FUNCTION "ROLL_PB21" : Void
{ S7_Optimized_Access := 'TRUE' }
VERSION : 0.1
VAR_TEMP
    r : Bool;
    a1 : Word;
    a2 : Word;
    activeDataBlock : Int;
    comparisonResults : Array[0..0] of Bool;
END_VAR
BEGIN
    #r := FALSE;
    #a1 := W#16#0000;
    #a2 := W#16#0000;
    #activeDataBlock := 0;
    // PB21, STEP 5 network 1
    #activeDataBlock := 15;
    // PB21, STEP 5 network 2
    #r := ((NOT "ROLL_IO".Input[3, 6]) AND (NOT "ROLL_State".M[13, 1]) AND (NOT "ROLL_State".M[5, 6]));
    "ROLL_State".M[99, 7] := #r;
    // PB21, STEP 5 network 3
    #r := ((NOT "ROLL_State".M[13, 3]) AND (NOT "ROLL_State".M[16, 6]) AND (NOT "ROLL_State".M[6, 0]) AND (NOT "ROLL_State".M[6, 2]) AND "ROLL_IO".Input[3, 0] AND "ROLL_IO".Input[5, 0] AND "ROLL_IO".Input[5, 2] AND "ROLL_IO".Input[5, 4]);
    "ROLL_State".M[100, 0] := #r;
    // PB21, STEP 5 network 4
    #r := "ROLL_State".M[190, 6];
    IF #r THEN "ROLL_State".M[100, 1] := TRUE; END_IF;
    #r := (((NOT "ROLL_State".M[190, 6]) AND "ROLL_IO".Input[5, 3]) OR (NOT "ROLL_IO".Input[0, 1]) OR (NOT "ROLL_State".M[0, 3]) OR (NOT "ROLL_State".M[100, 0]) OR "ROLL_State".M[190, 5]);
    IF #r THEN "ROLL_State".M[100, 1] := FALSE; END_IF;
    // PB21, STEP 5 network 5
    #r := "ROLL_State".M[190, 6];
    IF #r THEN "ROLL_State".M[100, 2] := TRUE; END_IF;
    #r := (("ROLL_IO".Input[5, 3] AND "ROLL_IO".Input[5, 6]) OR (NOT "ROLL_IO".Input[0, 1]) OR (NOT "ROLL_State".M[0, 3]) OR (NOT "ROLL_State".M[100, 0]) OR "ROLL_State".M[190, 5]);
    IF #r THEN "ROLL_State".M[100, 2] := FALSE; END_IF;
    // PB21, STEP 5 network 6
    #r := "ROLL_State".M[190, 6];
    IF #r THEN "ROLL_State".M[100, 3] := TRUE; END_IF;
    #r := (((NOT "ROLL_IO".Input[7, 5]) AND (NOT "ROLL_State".M[190, 6])) OR (NOT "ROLL_IO".Input[0, 1]) OR (NOT "ROLL_State".M[0, 3]) OR (NOT "ROLL_State".M[100, 0]) OR "ROLL_State".M[190, 5] OR "ROLL_State".M[5, 6] OR "ROLL_State".M[8, 5]);
    IF #r THEN "ROLL_State".M[100, 3] := FALSE; END_IF;
    // PB21, STEP 5 network 7
    #r := "ROLL_State".M[190, 6];
    IF #r THEN "ROLL_State".M[100, 4] := TRUE; END_IF;
    #r := (((NOT "ROLL_State".M[100, 0]) AND (NOT "ROLL_State".M[190, 6])) OR (NOT "ROLL_IO".Input[0, 1]) OR (NOT "ROLL_State".M[0, 3]) OR (NOT "ROLL_State".M[99, 7]) OR "ROLL_State".M[190, 5]);
    IF #r THEN "ROLL_State".M[100, 4] := FALSE; END_IF;
    // PB21, STEP 5 network 8
    #r := ((NOT "ROLL_State".M[31, 5]) AND (NOT "ROLL_State".M[5, 6]) AND ((NOT "ROLL_IO".Input[5, 6]) OR (NOT "ROLL_State".S5Timers[70].Q)) AND "ROLL_IO".Input[0, 2] AND "ROLL_IO".Input[3, 1] AND "ROLL_State".M[100, 0]);
    "ROLL_State".M[100, 5] := #r;
    // PB21, STEP 5 network 9
    #r := ((("ROLL_IO".Input[7, 5] AND "ROLL_State".S5Timers[97].Q) OR (NOT "ROLL_State".S5Timers[96].Q)) AND "ROLL_State".M[0, 3] AND "ROLL_State".M[100, 5]);
    "ROLL_State".M[100, 6] := #r;
    // PB21, STEP 5 network 10
    #r := ((((NOT "ROLL_IO".Input[7, 5]) AND "ROLL_State".S5Timers[96].Q) OR (NOT "ROLL_State".S5Timers[97].Q)) AND "ROLL_State".M[0, 3] AND "ROLL_State".M[100, 5]);
    "ROLL_State".M[100, 7] := #r;
    // PB21, STEP 5 network 11
    #r := "ROLL_State".M[190, 6];
    IF #r THEN "ROLL_State".M[101, 1] := TRUE; END_IF;
    #r := (((NOT "ROLL_State".M[190, 6]) AND "ROLL_IO".Input[5, 3] AND "ROLL_IO".Input[5, 6] AND "ROLL_IO".Input[6, 0]) OR (NOT "ROLL_IO".Input[0, 1]) OR (NOT "ROLL_State".M[0, 3]) OR (NOT "ROLL_State".M[100, 0]) OR "ROLL_State".M[190, 5]);
    IF #r THEN "ROLL_State".M[101, 1] := FALSE; END_IF;
    // PB21, STEP 5 network 12
    #r := "ROLL_State".M[190, 6];
    IF #r THEN "ROLL_State".M[101, 2] := TRUE; END_IF;
    #r := (((NOT "ROLL_State".M[190, 6]) AND "ROLL_IO".Input[5, 3] AND "ROLL_IO".Input[5, 6] AND "ROLL_IO".Input[6, 0]) OR (NOT "ROLL_IO".Input[0, 1]) OR (NOT "ROLL_State".M[0, 3]) OR (NOT "ROLL_State".M[100, 0]) OR "ROLL_State".M[190, 5]);
    IF #r THEN "ROLL_State".M[101, 2] := FALSE; END_IF;
    // PB21, STEP 5 network 13
    #r := "ROLL_State".M[190, 6];
    IF #r THEN "ROLL_State".M[101, 3] := TRUE; END_IF;
    #r := (((NOT "ROLL_State".M[190, 6]) AND ((NOT "ROLL_IO".Input[7, 5]) OR "ROLL_IO".Input[6, 0])) OR (NOT "ROLL_IO".Input[0, 1]) OR (NOT "ROLL_State".M[0, 3]) OR (NOT "ROLL_State".M[100, 0]) OR "ROLL_State".M[190, 5] OR "ROLL_State".M[5, 6] OR "ROLL_State".M[8, 5]);
    IF #r THEN "ROLL_State".M[101, 3] := FALSE; END_IF;
    // PB21, STEP 5 network 14
    #r := "ROLL_State".M[190, 6];
    IF #r THEN "ROLL_State".M[101, 4] := TRUE; END_IF;
    #r := (((NOT "ROLL_State".M[190, 6]) AND "ROLL_IO".Input[6, 0]) OR (NOT "ROLL_IO".Input[0, 1]) OR (NOT "ROLL_State".M[0, 3]) OR (NOT "ROLL_State".M[100, 0]) OR (NOT "ROLL_State".M[99, 7]) OR "ROLL_State".M[190, 5]);
    IF #r THEN "ROLL_State".M[101, 4] := FALSE; END_IF;
    // PB21, STEP 5 network 15
    #a2 := #a1;
    #a1 := W#16#2005;
    #r := "ROLL_IO".Input[6, 0];
    "ROLL_TimerOp"(Number := 121, Operation := 0, Signal := #r, Preset := #a1);
    // PB21, STEP 5 network 16
    #r := ((NOT "ROLL_State".M[31, 5]) AND (NOT "ROLL_State".M[5, 6]) AND (((NOT "ROLL_State".S5Timers[121].Q) AND "ROLL_State".M[101, 5]) OR (NOT "ROLL_IO".Input[6, 0])) AND "ROLL_IO".Input[0, 2] AND "ROLL_IO".Input[3, 1] AND "ROLL_State".M[100, 0]);
    "ROLL_State".M[101, 5] := #r;
    // PB21, STEP 5 network 17
    #r := ((("ROLL_IO".Input[7, 5] AND "ROLL_State".S5Timers[97].Q) OR (NOT "ROLL_State".S5Timers[96].Q)) AND "ROLL_State".M[101, 5]);
    "ROLL_State".M[101, 6] := #r;
    // PB21, STEP 5 network 18
    #r := ((((NOT "ROLL_IO".Input[7, 5]) AND "ROLL_State".S5Timers[96].Q) OR (NOT "ROLL_State".S5Timers[97].Q)) AND "ROLL_State".M[101, 5]);
    "ROLL_State".M[101, 7] := #r;
    // PB21, STEP 5 network 19
    #r := "ROLL_State".M[190, 6];
    IF #r THEN "ROLL_State".M[102, 1] := TRUE; END_IF;
    #r := (((NOT "ROLL_State".M[190, 6]) AND "ROLL_IO".Input[5, 3] AND "ROLL_IO".Input[5, 6] AND "ROLL_IO".Input[6, 0] AND "ROLL_IO".Input[6, 2]) OR (NOT "ROLL_IO".Input[0, 1]) OR (NOT "ROLL_State".M[0, 3]) OR (NOT "ROLL_State".M[100, 0]) OR "ROLL_State".M[190, 5]);
    IF #r THEN "ROLL_State".M[102, 1] := FALSE; END_IF;
    // PB21, STEP 5 network 20
    #r := "ROLL_State".M[190, 6];
    IF #r THEN "ROLL_State".M[102, 2] := TRUE; END_IF;
    #r := (((NOT "ROLL_State".M[190, 6]) AND "ROLL_IO".Input[6, 2]) OR (NOT "ROLL_IO".Input[0, 1]) OR (NOT "ROLL_State".M[0, 3]) OR (NOT "ROLL_State".M[100, 0]) OR "ROLL_State".M[190, 5]);
    IF #r THEN "ROLL_State".M[102, 2] := FALSE; END_IF;
    // PB21, STEP 5 network 21
    #r := "ROLL_State".M[190, 6];
    IF #r THEN "ROLL_State".M[102, 3] := TRUE; END_IF;
    #r := (((NOT "ROLL_State".M[190, 6]) AND ((NOT "ROLL_IO".Input[7, 5]) OR "ROLL_IO".Input[6, 2])) OR (NOT "ROLL_IO".Input[0, 1]) OR (NOT "ROLL_State".M[0, 3]) OR (NOT "ROLL_State".M[100, 0]) OR "ROLL_State".M[190, 5] OR "ROLL_State".M[5, 6] OR "ROLL_State".M[8, 5]);
    IF #r THEN "ROLL_State".M[102, 3] := FALSE; END_IF;
    // PB21, STEP 5 network 22
    #r := "ROLL_State".M[190, 6];
    IF #r THEN "ROLL_State".M[102, 4] := TRUE; END_IF;
    #r := (((NOT "ROLL_State".M[190, 6]) AND "ROLL_IO".Input[6, 2]) OR (NOT "ROLL_IO".Input[0, 1]) OR (NOT "ROLL_State".M[0, 3]) OR (NOT "ROLL_State".M[100, 0]) OR (NOT "ROLL_State".M[99, 7]) OR "ROLL_State".M[190, 5]);
    IF #r THEN "ROLL_State".M[102, 4] := FALSE; END_IF;
    // PB21, STEP 5 network 23
    #r := ((NOT "ROLL_State".M[31, 5]) AND (NOT "ROLL_State".M[5, 6]) AND (NOT "ROLL_State".S5Timers[72].Q) AND "ROLL_IO".Input[0, 2] AND "ROLL_IO".Input[3, 1] AND "ROLL_State".M[100, 0]);
    "ROLL_State".M[102, 5] := #r;
    // PB21, STEP 5 network 24
    #r := ((("ROLL_IO".Input[7, 5] AND "ROLL_State".S5Timers[97].Q) OR (NOT "ROLL_State".S5Timers[96].Q)) AND "ROLL_State".M[0, 3] AND "ROLL_State".M[102, 5]);
    "ROLL_State".M[102, 6] := #r;
    // PB21, STEP 5 network 25
    #r := ((((NOT "ROLL_IO".Input[7, 5]) AND "ROLL_State".S5Timers[96].Q) OR (NOT "ROLL_State".S5Timers[97].Q) OR "ROLL_State".M[0, 4]) AND "ROLL_State".M[102, 5]);
    "ROLL_State".M[102, 7] := #r;
    // PB21, STEP 5 network 26
    #r := "ROLL_State".M[190, 6];
    IF #r THEN "ROLL_State".M[105, 1] := TRUE; END_IF;
    #r := (((NOT "ROLL_State".M[190, 6]) AND "ROLL_State".M[0, 4]) OR (NOT "ROLL_IO".Input[0, 1]) OR (NOT "ROLL_State".M[0, 3]) OR (NOT "ROLL_State".M[100, 0]) OR "ROLL_State".M[190, 5]);
    IF #r THEN "ROLL_State".M[105, 1] := FALSE; END_IF;
    // PB21, STEP 5 network 27
    #r := "ROLL_State".M[190, 6];
    IF #r THEN "ROLL_State".M[105, 2] := TRUE; END_IF;
    #r := ((NOT "ROLL_IO".Input[0, 1]) OR (NOT "ROLL_State".M[0, 3]) OR (NOT "ROLL_State".M[100, 0]) OR "ROLL_IO".Input[6, 2] OR "ROLL_State".M[190, 5]);
    IF #r THEN "ROLL_State".M[105, 2] := FALSE; END_IF;
    // PB21, STEP 5 network 28
    #r := "ROLL_State".M[190, 6];
    IF #r THEN "ROLL_State".M[105, 3] := TRUE; END_IF;
    #r := (((NOT "ROLL_State".M[190, 6]) AND ((NOT "ROLL_IO".Input[7, 5]) OR "ROLL_State".M[0, 4])) OR (NOT "ROLL_IO".Input[0, 1]) OR (NOT "ROLL_State".M[0, 3]) OR (NOT "ROLL_State".M[100, 0]) OR "ROLL_State".M[190, 5] OR "ROLL_State".M[5, 6] OR "ROLL_State".M[8, 5]);
    IF #r THEN "ROLL_State".M[105, 3] := FALSE; END_IF;
    // PB21, STEP 5 network 29
    #r := "ROLL_State".M[190, 6];
    IF #r THEN "ROLL_State".M[105, 4] := TRUE; END_IF;
    #r := (((NOT "ROLL_State".M[190, 6]) AND "ROLL_State".M[0, 4]) OR (NOT "ROLL_IO".Input[0, 1]) OR (NOT "ROLL_State".M[0, 3]) OR (NOT "ROLL_State".M[100, 0]) OR (NOT "ROLL_State".M[99, 7]) OR "ROLL_State".M[190, 5]);
    IF #r THEN "ROLL_State".M[105, 4] := FALSE; END_IF;
    // PB21, STEP 5 network 30
    #a2 := #a1;
    #a1 := W#16#2005;
    #r := "ROLL_State".M[0, 4];
    "ROLL_TimerOp"(Number := 120, Operation := 0, Signal := #r, Preset := #a1);
    // PB21, STEP 5 network 31
    #r := ((NOT "ROLL_State".M[31, 5]) AND (NOT "ROLL_State".M[5, 6]) AND (((NOT "ROLL_State".S5Timers[120].Q) AND "ROLL_State".M[105, 5]) OR (NOT "ROLL_State".M[0, 4])) AND "ROLL_IO".Input[0, 2] AND "ROLL_IO".Input[3, 1] AND "ROLL_State".M[100, 0]);
    "ROLL_State".M[105, 5] := #r;
    // PB21, STEP 5 network 32
    #r := ((("ROLL_IO".Input[7, 5] AND "ROLL_State".S5Timers[97].Q) OR (NOT "ROLL_State".S5Timers[96].Q)) AND "ROLL_State".M[105, 5]);
    "ROLL_State".M[105, 6] := #r;
    // PB21, STEP 5 network 33
    #r := ((((NOT "ROLL_IO".Input[7, 5]) AND "ROLL_State".S5Timers[96].Q) OR (NOT "ROLL_State".S5Timers[97].Q)) AND "ROLL_State".M[105, 5]);
    "ROLL_State".M[105, 7] := #r;
    // PB21, STEP 5 network 34
    #r := ((((NOT "ROLL_IO".Input[5, 5]) AND ("ROLL_State".M[40, 5] OR "ROLL_State".M[42, 1]) AND "ROLL_State".M[31, 5]) OR (NOT "ROLL_IO".Input[5, 6])) AND "ROLL_IO".Input[0, 2] AND "ROLL_IO".Input[3, 1] AND "ROLL_State".M[100, 0]);
    "ROLL_State".M[103, 0] := #r;
    // PB21, STEP 5 network 35
    #r := (((NOT "ROLL_IO".Input[5, 3]) OR (NOT "ROLL_IO".Input[6, 0]) OR (NOT "ROLL_State".S5Timers[121].Q)) AND "ROLL_IO".Input[3, 1] AND "ROLL_State".M[100, 0] AND "ROLL_State".M[31, 5]);
    "ROLL_State".M[103, 3] := #r;
    // PB21, STEP 5 network 36
    #r := (((NOT "ROLL_IO".Input[5, 6]) AND "ROLL_IO".Input[0, 2]) OR (("ROLL_State".M[103, 0] OR "ROLL_State".M[103, 3]) AND "ROLL_State".S5Timers[62].Q AND "ROLL_State".S5Timers[97].Q));
    "ROLL_State".M[103, 1] := #r;
    // PB21, STEP 5 network 37
    #r := ((NOT "ROLL_IO".Input[6, 2]) AND "ROLL_IO".Input[3, 1] AND "ROLL_State".M[100, 0] AND "ROLL_State".M[31, 5]);
    "ROLL_State".M[103, 4] := #r;
    // PB21, STEP 5 network 38
    #a2 := #a1;
    #a1 := W#16#1050;
    #r := ("ROLL_IO".Output[22, 3] AND "ROLL_State".M[103, 4]);
    "ROLL_TimerOp"(Number := 119, Operation := 1, Signal := #r, Preset := #a1);
    // PB21, STEP 5 network 39
    #r := (((("ROLL_State".M[103, 0] OR "ROLL_State".M[103, 3]) AND "ROLL_State".S5Timers[96].Q) OR "ROLL_State".M[103, 4] OR "ROLL_State".S5Timers[119].Q) AND "ROLL_State".S5Timers[62].Q);
    "ROLL_State".M[103, 2] := #r;
    // PB21, STEP 5 network 40
    #r := "ROLL_State".M[190, 6];
    IF #r THEN "ROLL_State".M[104, 0] := TRUE; END_IF;
    #r := (((NOT "ROLL_State".M[190, 6]) AND ((NOT "ROLL_IO".Input[5, 0]) OR (NOT "ROLL_IO".Input[5, 2]) OR (NOT "ROLL_IO".Input[5, 4]))) OR (NOT "ROLL_IO".Input[0, 1]) OR (NOT "ROLL_IO".Input[7, 0]) OR (NOT "ROLL_State".M[26, 5]) OR (NOT "ROLL_State".M[99, 7]) OR "ROLL_State".M[16, 6] OR "ROLL_State".M[190, 5]);
    IF #r THEN "ROLL_State".M[104, 0] := FALSE; END_IF;
    // PB21, STEP 5 network 41
    #r := "ROLL_State".M[190, 6];
    IF #r THEN "ROLL_State".M[104, 1] := TRUE; END_IF;
    #r := (((NOT "ROLL_State".M[190, 6]) AND ((NOT "ROLL_IO".Input[5, 0]) OR (NOT "ROLL_IO".Input[5, 2]) OR (NOT "ROLL_IO".Input[5, 4]))) OR (NOT "ROLL_IO".Input[0, 1]) OR (NOT "ROLL_State".M[26, 0]) OR (NOT "ROLL_State".M[99, 7]) OR "ROLL_State".M[16, 6] OR "ROLL_State".M[190, 5]);
    IF #r THEN "ROLL_State".M[104, 1] := FALSE; END_IF;
    // PB21, STEP 5 network 42
    #r := "ROLL_State".M[190, 6];
    IF #r THEN "ROLL_State".M[104, 4] := TRUE; END_IF;
    #r := (((NOT "ROLL_State".M[190, 6]) AND ((NOT "ROLL_IO".Input[5, 0]) OR (NOT "ROLL_IO".Input[5, 2]) OR (NOT "ROLL_IO".Input[5, 4]))) OR (NOT "ROLL_IO".Input[0, 1]) OR (NOT "ROLL_IO".Input[4, 7]) OR (NOT "ROLL_State".M[27, 4]) OR (NOT "ROLL_State".M[99, 7]) OR "ROLL_State".M[16, 6] OR "ROLL_State".M[190, 5]);
    IF #r THEN "ROLL_State".M[104, 4] := FALSE; END_IF;
    // PB21, STEP 5 network 43
    #r := "ROLL_State".M[190, 6];
    IF #r THEN "ROLL_State".M[104, 5] := TRUE; END_IF;
    #r := (((NOT "ROLL_State".M[190, 6]) AND "ROLL_IO".Input[5, 3] AND "ROLL_IO".Input[5, 6] AND "ROLL_IO".Input[6, 0] AND "ROLL_IO".Input[6, 2]) OR (NOT "ROLL_IO".Input[0, 1]) OR (NOT "ROLL_State".M[100, 0]) OR (NOT "ROLL_State".M[24, 1]) OR "ROLL_State".M[190, 5]);
    IF #r THEN "ROLL_State".M[104, 5] := FALSE; END_IF;
    // PB21, STEP 5 network 44
    #r := "ROLL_State".M[190, 6];
    IF #r THEN "ROLL_State".M[104, 6] := TRUE; END_IF;
    #r := (((NOT "ROLL_State".M[190, 6]) AND (("ROLL_IO".Input[5, 3] AND "ROLL_IO".Input[5, 6] AND "ROLL_IO".Input[6, 0]) OR (NOT "ROLL_IO".Input[7, 5]))) OR (NOT "ROLL_IO".Input[0, 1]) OR (NOT "ROLL_State".M[100, 0]) OR (NOT "ROLL_State".M[25, 0]) OR "ROLL_State".M[190, 5] OR "ROLL_State".M[5, 6] OR "ROLL_State".M[8, 5]);
    IF #r THEN "ROLL_State".M[104, 6] := FALSE; END_IF;
    // PB21, STEP 5 network 45
    #r := "ROLL_State".S5Timers[59].Q;
    "ROLL_IO".Output[17, 0] := #r;
    // PB21, STEP 5 network 46
    #r := ("ROLL_IO".Input[6, 5] AND "ROLL_State".M[100, 0]);
    "ROLL_IO".Output[17, 5] := #r;
    RETURN;
END_FUNCTION

FUNCTION "ROLL_PB23" : Void
{ S7_Optimized_Access := 'TRUE' }
VERSION : 0.1
VAR_TEMP
    r : Bool;
    a1 : Word;
    a2 : Word;
    activeDataBlock : Int;
    comparisonResults : Array[0..0] of Bool;
END_VAR
BEGIN
    #r := FALSE;
    #a1 := W#16#0000;
    #a2 := W#16#0000;
    #activeDataBlock := 0;
    // PB23, STEP 5 network 1
    #activeDataBlock := 15;
    // PB23, STEP 5 network 2
    #r := (("ROLL_State".M[40, 3] OR "ROLL_State".M[40, 4] OR "ROLL_State".M[40, 5]) AND "ROLL_State".M[111, 4]);
    "ROLL_State".M[240, 0] := #r;
    // PB23, STEP 5 network 3
    #a2 := #a1;
    #a1 := W#16#2120;
    #r := "ROLL_State".M[240, 0];
    "ROLL_TimerOp"(Number := 51, Operation := 1, Signal := #r, Preset := #a1);
    #r := "ROLL_State".S5Timers[51].Q;
    "ROLL_IO".Output[19, 0] := #r;
    // PB23, STEP 5 network 4
    #a2 := #a1;
    #a1 := W#16#1050;
    #r := ((NOT "ROLL_State".M[6, 1]) AND ("ROLL_State".M[40, 4] OR "ROLL_State".M[40, 5]) AND "ROLL_IO".Output[19, 0] AND "ROLL_State".M[240, 0] AND "ROLL_State".M[35, 2] AND "ROLL_State".S5Timers[70].Q);
    "ROLL_TimerOp"(Number := 52, Operation := 0, Signal := #r, Preset := #a1);
    #r := "ROLL_State".S5Timers[52].Q;
    "ROLL_IO".Output[19, 1] := #r;
    // PB23, STEP 5 network 5
    #r := ("ROLL_IO".Input[0, 2] AND "ROLL_IO".Input[0, 4]);
    IF #r THEN "ROLL_State".M[103, 7] := TRUE; END_IF;
    #r := (NOT "ROLL_State".S5Timers[59].Q);
    IF #r THEN "ROLL_State".M[103, 7] := FALSE; END_IF;
    // PB23, STEP 5 network 6
    #a2 := #a1;
    #a1 := W#16#3360;
    #r := "ROLL_State".S5Timers[59].Q;
    "ROLL_TimerOp"(Number := 76, Operation := 0, Signal := #r, Preset := #a1);
    // PB23, STEP 5 network 7
    #r := ((NOT "ROLL_State".M[13, 3]) AND (NOT "ROLL_State".M[5, 6]) AND (NOT "ROLL_State".M[6, 2]) AND (NOT "ROLL_State".M[6, 3]) AND (((NOT "ROLL_State".S5Timers[76].Q) AND "ROLL_IO".Input[2, 2]) OR "ROLL_State".M[103, 7] OR "ROLL_State".M[152, 0]) AND ("ROLL_IO".Input[2, 2] OR "ROLL_State".M[152, 0]) AND "ROLL_IO".Input[3, 4] AND "ROLL_IO".Input[5, 6] AND "ROLL_State".S5Timers[59].Q);
    "ROLL_IO".Output[19, 5] := #r;
    // PB23, STEP 5 network 8
    #r := ((NOT "ROLL_State".M[5, 6]) AND (NOT "ROLL_State".M[6, 1]) AND ("ROLL_IO".Input[0, 1] OR "ROLL_IO".Input[0, 2]) AND "ROLL_IO".Input[3, 1] AND "ROLL_IO".Input[3, 4] AND "ROLL_State".M[0, 3] AND "ROLL_State".M[100, 0] AND "ROLL_State".S5Timers[70].Q);
    "ROLL_State".M[240, 0] := #r;
    // PB23, STEP 5 network 9
    #r := ((NOT "ROLL_IO".Output[20, 6]) AND (NOT "ROLL_State".M[5, 6]) AND (NOT "ROLL_State".M[8, 5]) AND (NOT "ROLL_State".S5Timers[96].Q) AND (("ROLL_State".M[100, 0] AND "ROLL_State".M[103, 1]) OR "ROLL_State".M[102, 6] OR "ROLL_State".M[104, 6]));
    "ROLL_IO".Output[20, 4] := #r;
    "ROLL_IO".Output[22, 6] := #r;
    // PB23, STEP 5 network 10
    #r := ((NOT "ROLL_IO".Output[20, 1]) AND ("ROLL_State".M[104, 0] OR "ROLL_State".M[104, 1] OR "ROLL_State".M[104, 4] OR "ROLL_State".M[152, 1]) AND "ROLL_State".M[99, 7]);
    "ROLL_IO".Output[20, 6] := #r;
    // PB23, STEP 5 network 11
    #r := ("ROLL_State".M[102, 7] OR "ROLL_State".M[103, 2] OR "ROLL_State".M[104, 5]);
    "ROLL_State".M[240, 0] := #r;
    // PB23, STEP 5 network 12
    #r := ((NOT "ROLL_State".M[13, 4]) AND (NOT "ROLL_State".M[6, 0]) AND (NOT "ROLL_State".M[6, 2]) AND (NOT "ROLL_State".M[7, 7]) AND "ROLL_IO".Input[3, 1] AND "ROLL_IO".Input[5, 0] AND "ROLL_IO".Input[5, 2] AND "ROLL_IO".Input[5, 4] AND "ROLL_State".M[240, 0]);
    "ROLL_IO".Output[20, 1] := #r;
    // PB23, STEP 5 network 13
    #r := "ROLL_State".M[103, 1];
    "ROLL_IO".Output[22, 2] := #r;
    // PB23, STEP 5 network 14
    #r := ("ROLL_State".M[102, 1] OR "ROLL_State".M[102, 2] OR "ROLL_State".M[102, 3] OR "ROLL_State".M[102, 6] OR "ROLL_State".M[102, 7] OR "ROLL_State".M[103, 2]);
    "ROLL_IO".Output[22, 3] := #r;
    // PB23, STEP 5 network 15
    #r := "ROLL_State".S5Timers[85].Q;
    "ROLL_IO".Output[21, 3] := #r;
    // PB23, STEP 5 network 16
    #a2 := #a1;
    #a1 := W#16#1020;
    #r := "ROLL_IO".Output[20, 6];
    "ROLL_TimerOp"(Number := 47, Operation := 1, Signal := #r, Preset := #a1);
    // PB23, STEP 5 network 17
    #r := ((NOT "ROLL_IO".Output[21, 5]) AND (NOT "ROLL_IO".Output[22, 3]) AND (NOT "ROLL_IO".Output[22, 6]) AND (("ROLL_IO".Output[21, 4] AND "ROLL_State".S5Timers[47].Q) OR "ROLL_State".M[104, 0] OR "ROLL_State".M[152, 1]));
    "ROLL_IO".Output[21, 4] := #r;
    // PB23, STEP 5 network 18
    #r := ((NOT "ROLL_IO".Output[21, 4]) AND "ROLL_State".M[152, 0]);
    "ROLL_IO".Output[21, 5] := #r;
    // PB23, STEP 5 network 19
    RETURN;
END_FUNCTION

FUNCTION "ROLL_PB24" : Void
{ S7_Optimized_Access := 'TRUE' }
VERSION : 0.1
VAR_TEMP
    r : Bool;
    a1 : Word;
    a2 : Word;
    activeDataBlock : Int;
    comparisonResults : Array[0..0] of Bool;
END_VAR
BEGIN
    #r := FALSE;
    #a1 := W#16#0000;
    #a2 := W#16#0000;
    #activeDataBlock := 0;
    // PB24, STEP 5 network 1
    #activeDataBlock := 15;
    // PB24, STEP 5 network 2
    #r := ("ROLL_IO".Input[5, 0] AND "ROLL_State".M[13, 3] AND "ROLL_State".S5Timers[59].Q);
    "ROLL_State".M[240, 0] := #r;
    // PB24, STEP 5 network 3
    #a2 := #a1;
    #a1 := "ROLL_GetDW"(DbNumber := #activeDataBlock, Index := 54);
    #r := (NOT "ROLL_State".S5Timers[53].Q);
    "ROLL_TimerOp"(Number := 54, Operation := 0, Signal := #r, Preset := #a1);
    #a2 := #a1;
    #a1 := "ROLL_GetDW"(DbNumber := #activeDataBlock, Index := 53);
    #r := "ROLL_State".S5Timers[54].Q;
    "ROLL_TimerOp"(Number := 53, Operation := 1, Signal := #r, Preset := #a1);
    #r := "ROLL_State".M[240, 0];
    "ROLL_TimerOp"(Number := 53, Operation := 2, Signal := #r, Preset := #a1);
    #r := ((NOT "ROLL_State".M[40, 5]) AND "ROLL_State".S5Timers[53].Q);
    "ROLL_IO".Output[19, 4] := #r;
    // PB24, STEP 5 network 4
    RETURN;
END_FUNCTION

FUNCTION "ROLL_PB25" : Void
{ S7_Optimized_Access := 'TRUE' }
VERSION : 0.1
VAR_TEMP
    r : Bool;
    a1 : Word;
    a2 : Word;
    activeDataBlock : Int;
    comparisonResults : Array[0..14] of Bool;
END_VAR
BEGIN
    #r := FALSE;
    #a1 := W#16#0000;
    #a2 := W#16#0000;
    #activeDataBlock := 0;
    // PB25, STEP 5 network 1
    #activeDataBlock := 15;
    // PB25, STEP 5 network 2
    #a2 := #a1;
    #a1 := "ROLL_GetM"(FirstByte := 5, Width := 8);
    #a2 := #a1;
    #a1 := W#16#0000;
    #comparisonResults[0] := (WORD_TO_INT(#a2) <> WORD_TO_INT(#a1));
    #r := #comparisonResults[0];
    "ROLL_State".M[87, 0] := #r;
    // PB25, STEP 5 network 3
    #a2 := #a1;
    #a1 := "ROLL_GetM"(FirstByte := 6, Width := 8);
    #a2 := #a1;
    #a1 := W#16#0000;
    #comparisonResults[1] := (WORD_TO_INT(#a2) <> WORD_TO_INT(#a1));
    #r := #comparisonResults[1];
    "ROLL_State".M[87, 1] := #r;
    // PB25, STEP 5 network 4
    #a2 := #a1;
    #a1 := "ROLL_GetM"(FirstByte := 7, Width := 8);
    #a2 := #a1;
    #a1 := W#16#0000;
    #comparisonResults[2] := (WORD_TO_INT(#a2) <> WORD_TO_INT(#a1));
    #r := #comparisonResults[2];
    "ROLL_State".M[87, 2] := #r;
    // PB25, STEP 5 network 5
    #a2 := #a1;
    #a1 := "ROLL_GetM"(FirstByte := 8, Width := 8);
    #a2 := #a1;
    #a1 := W#16#0000;
    #comparisonResults[3] := (WORD_TO_INT(#a2) <> WORD_TO_INT(#a1));
    #r := #comparisonResults[3];
    "ROLL_State".M[87, 3] := #r;
    // PB25, STEP 5 network 6
    #a2 := #a1;
    #a1 := "ROLL_GetM"(FirstByte := 9, Width := 8);
    #a2 := #a1;
    #a1 := W#16#0000;
    #comparisonResults[4] := (WORD_TO_INT(#a2) <> WORD_TO_INT(#a1));
    #r := #comparisonResults[4];
    "ROLL_State".M[87, 4] := #r;
    // PB25, STEP 5 network 7
    #a2 := #a1;
    #a1 := "ROLL_GetM"(FirstByte := 10, Width := 8);
    #a2 := #a1;
    #a1 := W#16#0000;
    #comparisonResults[5] := (WORD_TO_INT(#a2) <> WORD_TO_INT(#a1));
    #r := #comparisonResults[5];
    "ROLL_State".M[87, 5] := #r;
    // PB25, STEP 5 network 8
    #a2 := #a1;
    #a1 := "ROLL_GetM"(FirstByte := 11, Width := 8);
    #a2 := #a1;
    #a1 := W#16#0000;
    #comparisonResults[6] := (WORD_TO_INT(#a2) <> WORD_TO_INT(#a1));
    #r := #comparisonResults[6];
    "ROLL_State".M[87, 6] := #r;
    // PB25, STEP 5 network 9
    #a2 := #a1;
    #a1 := "ROLL_GetM"(FirstByte := 12, Width := 8);
    #a2 := #a1;
    #a1 := W#16#0000;
    #comparisonResults[7] := (WORD_TO_INT(#a2) <> WORD_TO_INT(#a1));
    #r := #comparisonResults[7];
    "ROLL_State".M[87, 7] := #r;
    // PB25, STEP 5 network 10
    #a2 := #a1;
    #a1 := "ROLL_GetM"(FirstByte := 13, Width := 8);
    #a2 := #a1;
    #a1 := W#16#0000;
    #comparisonResults[8] := (WORD_TO_INT(#a2) <> WORD_TO_INT(#a1));
    #r := #comparisonResults[8];
    "ROLL_State".M[88, 0] := #r;
    // PB25, STEP 5 network 11
    #a2 := #a1;
    #a1 := "ROLL_GetM"(FirstByte := 14, Width := 8);
    #a2 := #a1;
    #a1 := W#16#0000;
    #comparisonResults[9] := (WORD_TO_INT(#a2) <> WORD_TO_INT(#a1));
    #r := #comparisonResults[9];
    "ROLL_State".M[88, 1] := #r;
    // PB25, STEP 5 network 12
    #a2 := #a1;
    #a1 := "ROLL_GetM"(FirstByte := 15, Width := 8);
    #a2 := #a1;
    #a1 := W#16#0000;
    #comparisonResults[10] := (WORD_TO_INT(#a2) <> WORD_TO_INT(#a1));
    #r := #comparisonResults[10];
    "ROLL_State".M[88, 2] := #r;
    // PB25, STEP 5 network 13
    #a2 := #a1;
    #a1 := "ROLL_GetM"(FirstByte := 16, Width := 8);
    #a2 := #a1;
    #a1 := W#16#0000;
    #comparisonResults[11] := (WORD_TO_INT(#a2) <> WORD_TO_INT(#a1));
    #r := #comparisonResults[11];
    "ROLL_State".M[88, 3] := #r;
    // PB25, STEP 5 network 14
    #a2 := #a1;
    #a1 := "ROLL_GetM"(FirstByte := 17, Width := 8);
    #a2 := #a1;
    #a1 := W#16#0000;
    #comparisonResults[12] := (WORD_TO_INT(#a2) <> WORD_TO_INT(#a1));
    #r := #comparisonResults[12];
    "ROLL_State".M[88, 4] := #r;
    // PB25, STEP 5 network 15
    #a2 := #a1;
    #a1 := "ROLL_GetM"(FirstByte := 18, Width := 8);
    #a2 := #a1;
    #a1 := W#16#0000;
    #comparisonResults[13] := (WORD_TO_INT(#a2) <> WORD_TO_INT(#a1));
    #r := #comparisonResults[13];
    "ROLL_State".M[88, 5] := #r;
    // PB25, STEP 5 network 16
    #a2 := #a1;
    #a1 := "ROLL_GetM"(FirstByte := 19, Width := 8);
    #a2 := #a1;
    #a1 := W#16#0000;
    #comparisonResults[14] := (WORD_TO_INT(#a2) <> WORD_TO_INT(#a1));
    #r := #comparisonResults[14];
    "ROLL_State".M[88, 6] := #r;
    // PB25, STEP 5 network 17
    #r := ("ROLL_State".M[87, 0] OR "ROLL_State".M[87, 1] OR "ROLL_State".M[87, 2] OR "ROLL_State".M[87, 3] OR "ROLL_State".M[87, 4] OR "ROLL_State".M[87, 5] OR "ROLL_State".M[87, 6] OR "ROLL_State".M[87, 7] OR "ROLL_State".M[88, 0] OR "ROLL_State".M[88, 1] OR "ROLL_State".M[88, 2] OR "ROLL_State".M[88, 3] OR "ROLL_State".M[88, 4] OR "ROLL_State".M[88, 5] OR "ROLL_State".M[88, 6]);
    "ROLL_State".M[88, 7] := #r;
    // PB25, STEP 5 network 18
    #r := ("ROLL_IO".Input[1, 2] OR "ROLL_State".M[88, 7]);
    "ROLL_IO".Output[16, 4] := #r;
    // PB25, STEP 5 network 19
    #r := (("ROLL_State".M[3, 6] AND "ROLL_State".M[31, 6]) OR "ROLL_IO".Input[1, 2]);
    "ROLL_IO".Output[16, 5] := #r;
    // PB25, STEP 5 network 20
    #r := ("ROLL_IO".Input[1, 2] OR "ROLL_IO".Input[3, 4]);
    "ROLL_IO".Output[16, 0] := #r;
    // PB25, STEP 5 network 21
    #r := (((NOT "ROLL_State".M[31, 5]) AND "ROLL_State".M[28, 4]) OR ("ROLL_State".M[3, 6] AND "ROLL_State".M[74, 0]) OR "ROLL_IO".Input[1, 2]);
    "ROLL_IO".Output[16, 2] := #r;
    // PB25, STEP 5 network 22
    #r := (("ROLL_State".M[3, 6] AND "ROLL_State".M[31, 5]) OR "ROLL_IO".Input[1, 2] OR "ROLL_State".M[31, 4]);
    "ROLL_IO".Output[16, 3] := #r;
    // PB25, STEP 5 network 23
    #r := "ROLL_IO".Input[2, 0];
    "ROLL_IO".Output[19, 3] := #r;
    // PB25, STEP 5 network 24
    #r := (((("ROLL_IO".Input[14, 0] AND "ROLL_State".M[37, 1]) OR "ROLL_State".M[53, 6]) AND "ROLL_IO".Input[0, 2]) OR ("ROLL_IO".Input[0, 1] AND "ROLL_State".M[190, 6] AND "ROLL_State".M[20, 7]));
    IF #r THEN "ROLL_State".M[71, 5] := TRUE; END_IF;
    #r := (("ROLL_IO".Input[0, 1] AND "ROLL_State".M[190, 5] AND "ROLL_State".M[20, 7]) OR ("ROLL_IO".Input[0, 2] AND "ROLL_State".M[37, 2]));
    IF #r THEN "ROLL_State".M[71, 5] := FALSE; END_IF;
    #r := "ROLL_State".M[71, 5];
    "ROLL_IO".Output[17, 7] := #r;
    // PB25, STEP 5 network 25
    RETURN;
END_FUNCTION

FUNCTION "ROLL_PB50" : Void
{ S7_Optimized_Access := 'TRUE' }
VERSION : 0.1
VAR_TEMP
    r : Bool;
    a1 : Word;
    a2 : Word;
    activeDataBlock : Int;
    comparisonResults : Array[0..0] of Bool;
END_VAR
BEGIN
    #r := FALSE;
    #a1 := W#16#0000;
    #a2 := W#16#0000;
    #activeDataBlock := 0;
    // PB50, STEP 5 network 1
    #activeDataBlock := 15;
    // PB50, STEP 5 network 2
    #r := "ROLL_State".M[0, 1];
    IF #r THEN "ROLL_State".M[0, 2] := FALSE; END_IF;
    // PB50, STEP 5 network 3
    #a2 := #a1;
    #a1 := W#16#2008;
    #r := ((NOT "ROLL_State".M[0, 1]) AND "ROLL_IO".Input[3, 0]);
    "ROLL_TimerOp"(Number := 11, Operation := 0, Signal := #r, Preset := #a1);
    // PB50, STEP 5 network 4
    #a2 := #a1;
    #a1 := W#16#1020;
    #r := "ROLL_State".M[29, 0];
    "ROLL_TimerOp"(Number := 13, Operation := 0, Signal := #r, Preset := #a1);
    // PB50, STEP 5 network 5
    RETURN;
END_FUNCTION

FUNCTION "ROLL_PB51" : Void
{ S7_Optimized_Access := 'TRUE' }
VERSION : 0.1
VAR_TEMP
    r : Bool;
    a1 : Word;
    a2 : Word;
    activeDataBlock : Int;
    comparisonResults : Array[0..0] of Bool;
END_VAR
BEGIN
    #r := FALSE;
    #a1 := W#16#0000;
    #a2 := W#16#0000;
    #activeDataBlock := 0;
    // PB51, STEP 5 network 1
    #a2 := #a1;
    #a1 := W#16#2060;
    #r := "ROLL_IO".Output[24, 0];
    "ROLL_TimerOp"(Number := 15, Operation := 0, Signal := #r, Preset := #a1);
    // PB51, STEP 5 network 2
    #a2 := #a1;
    #a1 := W#16#3360;
    #r := ((NOT "ROLL_IO".Input[5, 6]) AND "ROLL_State".M[31, 5]);
    "ROLL_TimerOp"(Number := 16, Operation := 0, Signal := #r, Preset := #a1);
    // PB51, STEP 5 network 3
    #a2 := #a1;
    #a1 := W#16#1010;
    #r := "ROLL_State".M[37, 5];
    "ROLL_TimerOp"(Number := 18, Operation := 0, Signal := #r, Preset := #a1);
    // PB51, STEP 5 network 4
    #a2 := #a1;
    #a1 := W#16#2015;
    #r := (((NOT "ROLL_IO".Input[124, 1]) AND "ROLL_IO".Output[112, 1]) OR ((NOT "ROLL_IO".Input[124, 2]) AND "ROLL_IO".Output[112, 2]));
    "ROLL_TimerOp"(Number := 19, Operation := 0, Signal := #r, Preset := #a1);
    // PB51, STEP 5 network 5
    #a2 := #a1;
    #a1 := W#16#1010;
    #r := (("ROLL_IO".Input[123, 4] OR "ROLL_IO".Input[123, 5]) AND "ROLL_IO".Output[112, 0]);
    "ROLL_TimerOp"(Number := 20, Operation := 0, Signal := #r, Preset := #a1);
    // PB51, STEP 5 network 6
    #a2 := #a1;
    #a1 := W#16#1050;
    #r := "ROLL_IO".Input[123, 4];
    "ROLL_TimerOp"(Number := 21, Operation := 0, Signal := #r, Preset := #a1);
    // PB51, STEP 5 network 7
    #a2 := #a1;
    #a1 := W#16#2005;
    #r := ("ROLL_IO".Input[125, 0] AND "ROLL_IO".Input[125, 1]);
    "ROLL_TimerOp"(Number := 95, Operation := 0, Signal := #r, Preset := #a1);
    // PB51, STEP 5 network 8
    RETURN;
END_FUNCTION

FUNCTION "ROLL_PB52" : Void
{ S7_Optimized_Access := 'TRUE' }
VERSION : 0.1
VAR_TEMP
    r : Bool;
    a1 : Word;
    a2 : Word;
    activeDataBlock : Int;
    comparisonResults : Array[0..0] of Bool;
END_VAR
BEGIN
    #r := FALSE;
    #a1 := W#16#0000;
    #a2 := W#16#0000;
    #activeDataBlock := 0;
    // PB52, STEP 5 network 1
    #activeDataBlock := 15;
    // PB52, STEP 5 network 2
    #a2 := #a1;
    #a1 := "ROLL_GetDW"(DbNumber := #activeDataBlock, Index := 17);
    #r := ((NOT "ROLL_IO".Input[5, 5]) AND (NOT "ROLL_State".M[6, 3]) AND "ROLL_IO".Input[3, 1] AND "ROLL_State".M[4, 1] AND "ROLL_State".M[40, 5]);
    "ROLL_TimerOp"(Number := 17, Operation := 0, Signal := #r, Preset := #a1);
    // PB52, STEP 5 network 3
    #a2 := #a1;
    #a1 := "ROLL_GetDW"(DbNumber := #activeDataBlock, Index := 31);
    #r := ((NOT "ROLL_IO".Input[5, 3]) AND (NOT "ROLL_State".M[6, 1]) AND "ROLL_IO".Input[3, 1] AND "ROLL_State".M[4, 1]);
    "ROLL_TimerOp"(Number := 31, Operation := 0, Signal := #r, Preset := #a1);
    // PB52, STEP 5 network 4
    #a2 := #a1;
    #a1 := "ROLL_GetDW"(DbNumber := #activeDataBlock, Index := 32);
    #r := ((NOT "ROLL_IO".Input[6, 0]) AND (NOT "ROLL_State".M[6, 4]) AND "ROLL_IO".Input[3, 1] AND "ROLL_State".M[4, 1]);
    "ROLL_TimerOp"(Number := 32, Operation := 0, Signal := #r, Preset := #a1);
    // PB52, STEP 5 network 5
    #a2 := #a1;
    #a1 := "ROLL_GetDW"(DbNumber := #activeDataBlock, Index := 33);
    #r := ((NOT "ROLL_IO".Input[6, 2]) AND (NOT "ROLL_State".M[6, 5]) AND "ROLL_IO".Input[3, 1] AND "ROLL_State".M[4, 1]);
    "ROLL_TimerOp"(Number := 33, Operation := 0, Signal := #r, Preset := #a1);
    // PB52, STEP 5 network 6
    #a2 := #a1;
    #a1 := W#16#3030;
    #r := ((NOT "ROLL_State".M[0, 4]) AND (NOT "ROLL_State".M[6, 7]) AND "ROLL_IO".Input[3, 1] AND "ROLL_State".M[4, 1]);
    "ROLL_TimerOp"(Number := 35, Operation := 0, Signal := #r, Preset := #a1);
    // PB52, STEP 5 network 7
    #a2 := #a1;
    #a1 := W#16#3030;
    #r := ((NOT "ROLL_State".M[0, 4]) AND (NOT "ROLL_State".M[7, 0]) AND "ROLL_IO".Input[3, 1] AND "ROLL_State".M[4, 1]);
    "ROLL_TimerOp"(Number := 36, Operation := 0, Signal := #r, Preset := #a1);
    // PB52, STEP 5 network 8
    #a2 := #a1;
    #a1 := W#16#3030;
    #r := ((NOT "ROLL_State".M[0, 4]) AND (NOT "ROLL_State".M[7, 1]) AND "ROLL_IO".Input[3, 1] AND "ROLL_State".M[4, 1]);
    "ROLL_TimerOp"(Number := 37, Operation := 0, Signal := #r, Preset := #a1);
    // PB52, STEP 5 network 9
    #a2 := #a1;
    #a1 := W#16#3030;
    #r := ((NOT "ROLL_State".M[0, 4]) AND (NOT "ROLL_State".M[7, 2]) AND "ROLL_IO".Input[3, 1] AND "ROLL_State".M[4, 1]);
    "ROLL_TimerOp"(Number := 38, Operation := 0, Signal := #r, Preset := #a1);
    // PB52, STEP 5 network 10
    #a2 := #a1;
    #a1 := W#16#1005;
    #r := "ROLL_IO".Input[123, 1];
    "ROLL_TimerOp"(Number := 45, Operation := 0, Signal := #r, Preset := #a1);
    // PB52, STEP 5 network 11
    #a2 := #a1;
    #a1 := "ROLL_GetDW"(DbNumber := #activeDataBlock, Index := 58);
    #r := ("ROLL_IO".Input[3, 1] AND "ROLL_State".M[3, 6]);
    "ROLL_TimerOp"(Number := 58, Operation := 1, Signal := #r, Preset := #a1);
    #a2 := #a1;
    #a1 := "ROLL_GetDW"(DbNumber := #activeDataBlock, Index := 59);
    #r := ("ROLL_State".M[3, 6] AND "ROLL_State".S5Timers[58].Q);
    "ROLL_TimerOp"(Number := 59, Operation := 1, Signal := #r, Preset := #a1);
    // PB52, STEP 5 network 12
    #a2 := #a1;
    #a1 := "ROLL_GetDW"(DbNumber := #activeDataBlock, Index := 63);
    #r := (NOT "ROLL_State".S5Timers[62].Q);
    "ROLL_TimerOp"(Number := 63, Operation := 0, Signal := #r, Preset := #a1);
    #a2 := #a1;
    #a1 := "ROLL_GetDW"(DbNumber := #activeDataBlock, Index := 62);
    #r := "ROLL_State".S5Timers[63].Q;
    "ROLL_TimerOp"(Number := 62, Operation := 1, Signal := #r, Preset := #a1);
    #r := ((NOT "ROLL_State".M[103, 0]) AND (NOT "ROLL_State".M[103, 3]) AND (NOT "ROLL_State".M[103, 4]) AND (NOT "ROLL_State".S5Timers[119].Q));
    "ROLL_TimerOp"(Number := 62, Operation := 2, Signal := #r, Preset := #a1);
    // PB52, STEP 5 network 13
    #a2 := #a1;
    #a1 := W#16#2010;
    #r := "ROLL_IO".Input[5, 3];
    "ROLL_TimerOp"(Number := 70, Operation := 1, Signal := #r, Preset := #a1);
    // PB52, STEP 5 network 14
    #a2 := #a1;
    #a1 := W#16#2010;
    #r := "ROLL_IO".Input[6, 2];
    "ROLL_TimerOp"(Number := 72, Operation := 1, Signal := #r, Preset := #a1);
    // PB52, STEP 5 network 15
    #a2 := #a1;
    #a1 := "ROLL_GetDW"(DbNumber := #activeDataBlock, Index := 85);
    #r := "ROLL_State".M[41, 0];
    "ROLL_TimerOp"(Number := 85, Operation := 1, Signal := #r, Preset := #a1);
    // PB52, STEP 5 network 16
    RETURN;
END_FUNCTION

FUNCTION "ROLL_ReadInputs" : Void
{ S7_Optimized_Access := 'TRUE' }
VERSION : 0.1
VAR_TEMP
    b : Int;
    bit : Int;
END_VAR
BEGIN
    // Confirmed four-station profile: absent optional inputs are zero.
    FOR #b := 119 TO 125 DO
        FOR #bit := 0 TO 7 DO "ROLL_IO".Input[#b, #bit] := FALSE; END_FOR;
    END_FOR;
    IF "ROLL_IO".PhysicalIoConfigured AND NOT "ROLL_IO".Simulation THEN
        "ROLL_IO".Input[0, 0] := %I0.0;
        "ROLL_IO".Input[0, 1] := %I0.1;
        "ROLL_IO".Input[0, 2] := %I0.2;
        "ROLL_IO".Input[0, 3] := %I0.3;
        "ROLL_IO".Input[0, 4] := %I0.4;
        "ROLL_IO".Input[0, 5] := %I0.5;
        "ROLL_IO".Input[0, 6] := %I0.6;
        "ROLL_IO".Input[0, 7] := %I0.7;
        "ROLL_IO".Input[1, 0] := %I1.0;
        "ROLL_IO".Input[1, 1] := %I1.1;
        "ROLL_IO".Input[1, 2] := %I1.2;
        "ROLL_IO".Input[1, 3] := %I1.3;
        "ROLL_IO".Input[1, 4] := %I1.4;
        "ROLL_IO".Input[1, 5] := %I1.5;
        "ROLL_IO".Input[1, 6] := %I1.6;
        "ROLL_IO".Input[1, 7] := %I1.7;
        "ROLL_IO".Input[2, 0] := %I2.0;
        "ROLL_IO".Input[2, 1] := %I2.1;
        "ROLL_IO".Input[2, 2] := %I2.2;
        "ROLL_IO".Input[2, 3] := %I2.3;
        "ROLL_IO".Input[2, 4] := %I2.4;
        "ROLL_IO".Input[2, 5] := %I2.5;
        "ROLL_IO".Input[2, 6] := %I2.6;
        "ROLL_IO".Input[2, 7] := %I2.7;
        "ROLL_IO".Input[3, 0] := %I3.0;
        "ROLL_IO".Input[3, 1] := %I3.1;
        "ROLL_IO".Input[3, 2] := %I3.2;
        "ROLL_IO".Input[3, 3] := %I3.3;
        "ROLL_IO".Input[3, 4] := %I3.4;
        "ROLL_IO".Input[3, 5] := %I3.5;
        "ROLL_IO".Input[3, 6] := %I3.6;
        "ROLL_IO".Input[3, 7] := %I3.7;
        "ROLL_IO".Input[4, 0] := %I4.0;
        "ROLL_IO".Input[4, 1] := %I4.1;
        "ROLL_IO".Input[4, 2] := %I4.2;
        "ROLL_IO".Input[4, 3] := %I4.3;
        "ROLL_IO".Input[4, 4] := %I4.4;
        "ROLL_IO".Input[4, 5] := %I4.5;
        "ROLL_IO".Input[4, 6] := %I4.6;
        "ROLL_IO".Input[4, 7] := %I4.7;
        "ROLL_IO".Input[5, 0] := %I5.0;
        "ROLL_IO".Input[5, 1] := %I5.1;
        "ROLL_IO".Input[5, 2] := %I5.2;
        "ROLL_IO".Input[5, 3] := %I5.3;
        "ROLL_IO".Input[5, 4] := %I5.4;
        "ROLL_IO".Input[5, 5] := %I5.5;
        "ROLL_IO".Input[5, 6] := %I5.6;
        "ROLL_IO".Input[5, 7] := %I5.7;
        "ROLL_IO".Input[6, 0] := %I6.0;
        "ROLL_IO".Input[6, 1] := %I6.1;
        "ROLL_IO".Input[6, 2] := %I6.2;
        "ROLL_IO".Input[6, 3] := %I6.3;
        "ROLL_IO".Input[6, 4] := %I6.4;
        "ROLL_IO".Input[6, 5] := %I6.5;
        "ROLL_IO".Input[6, 6] := %I6.6;
        "ROLL_IO".Input[6, 7] := %I6.7;
        "ROLL_IO".Input[7, 0] := %I7.0;
        "ROLL_IO".Input[7, 1] := %I7.1;
        "ROLL_IO".Input[7, 2] := %I7.2;
        "ROLL_IO".Input[7, 3] := %I7.3;
        "ROLL_IO".Input[7, 4] := %I7.4;
        "ROLL_IO".Input[7, 5] := %I7.5;
        "ROLL_IO".Input[7, 6] := %I7.6;
        "ROLL_IO".Input[7, 7] := %I7.7;
        "ROLL_IO".Input[8, 0] := %I8.0;
        "ROLL_IO".Input[8, 1] := %I8.1;
        "ROLL_IO".Input[8, 2] := %I8.2;
        "ROLL_IO".Input[8, 3] := %I8.3;
        "ROLL_IO".Input[8, 4] := %I8.4;
        "ROLL_IO".Input[8, 5] := %I8.5;
        "ROLL_IO".Input[8, 6] := %I8.6;
        "ROLL_IO".Input[8, 7] := %I8.7;
        "ROLL_IO".Input[9, 0] := %I9.0;
        "ROLL_IO".Input[9, 1] := %I9.1;
        "ROLL_IO".Input[9, 2] := %I9.2;
        "ROLL_IO".Input[9, 3] := %I9.3;
        "ROLL_IO".Input[9, 4] := %I9.4;
        "ROLL_IO".Input[9, 5] := %I9.5;
        "ROLL_IO".Input[9, 6] := %I9.6;
        "ROLL_IO".Input[9, 7] := %I9.7;
        "ROLL_IO".Input[10, 0] := %I10.0;
        "ROLL_IO".Input[10, 1] := %I10.1;
        "ROLL_IO".Input[10, 2] := %I10.2;
        "ROLL_IO".Input[10, 3] := %I10.3;
        "ROLL_IO".Input[10, 4] := %I10.4;
        "ROLL_IO".Input[10, 5] := %I10.5;
        "ROLL_IO".Input[10, 6] := %I10.6;
        "ROLL_IO".Input[10, 7] := %I10.7;
        "ROLL_IO".Input[11, 0] := %I11.0;
        "ROLL_IO".Input[11, 1] := %I11.1;
        "ROLL_IO".Input[11, 2] := %I11.2;
        "ROLL_IO".Input[11, 3] := %I11.3;
        "ROLL_IO".Input[11, 4] := %I11.4;
        "ROLL_IO".Input[11, 5] := %I11.5;
        "ROLL_IO".Input[11, 6] := %I11.6;
        "ROLL_IO".Input[11, 7] := %I11.7;
        "ROLL_IO".Input[12, 0] := %I12.0;
        "ROLL_IO".Input[12, 1] := %I12.1;
        "ROLL_IO".Input[12, 2] := %I12.2;
        "ROLL_IO".Input[12, 3] := %I12.3;
        "ROLL_IO".Input[12, 4] := %I12.4;
        "ROLL_IO".Input[12, 5] := %I12.5;
        "ROLL_IO".Input[12, 6] := %I12.6;
        "ROLL_IO".Input[12, 7] := %I12.7;
        "ROLL_IO".Input[13, 0] := %I13.0;
        "ROLL_IO".Input[13, 1] := %I13.1;
        "ROLL_IO".Input[13, 2] := %I13.2;
        "ROLL_IO".Input[13, 3] := %I13.3;
        "ROLL_IO".Input[13, 4] := %I13.4;
        "ROLL_IO".Input[13, 5] := %I13.5;
        "ROLL_IO".Input[13, 6] := %I13.6;
        "ROLL_IO".Input[13, 7] := %I13.7;
        "ROLL_IO".Input[14, 0] := %I14.0;
        "ROLL_IO".Input[14, 1] := %I14.1;
        "ROLL_IO".Input[14, 2] := %I14.2;
        "ROLL_IO".Input[14, 3] := %I14.3;
        "ROLL_IO".Input[14, 4] := %I14.4;
        "ROLL_IO".Input[14, 5] := %I14.5;
        "ROLL_IO".Input[14, 6] := %I14.6;
        "ROLL_IO".Input[14, 7] := %I14.7;
        "ROLL_IO".Input[15, 0] := %I15.0;
        "ROLL_IO".Input[15, 1] := %I15.1;
        "ROLL_IO".Input[15, 2] := %I15.2;
        "ROLL_IO".Input[15, 3] := %I15.3;
        "ROLL_IO".Input[15, 4] := %I15.4;
        "ROLL_IO".Input[15, 5] := %I15.5;
        "ROLL_IO".Input[15, 6] := %I15.6;
        "ROLL_IO".Input[15, 7] := %I15.7;
    END_IF;
END_FUNCTION

FUNCTION "ROLL_WriteOutputs" : Void
{ S7_Optimized_Access := 'TRUE' }
VERSION : 0.1
VAR_TEMP
    enabled : Bool;
END_VAR
BEGIN
    IF "ROLL_IO".PhysicalIoConfigured THEN
        #enabled := "ROLL_IO".PhysicalOutputsEnabled AND NOT "ROLL_IO".Simulation AND NOT "ROLL_IO".ConversionFault;
        %Q16.0 := #enabled AND "ROLL_IO".Output[16, 0];
        %Q16.1 := #enabled AND "ROLL_IO".Output[16, 1];
        %Q16.2 := #enabled AND "ROLL_IO".Output[16, 2];
        %Q16.3 := #enabled AND "ROLL_IO".Output[16, 3];
        %Q16.4 := #enabled AND "ROLL_IO".Output[16, 4];
        %Q16.5 := #enabled AND "ROLL_IO".Output[16, 5];
        %Q16.6 := #enabled AND "ROLL_IO".Output[16, 6];
        %Q16.7 := #enabled AND "ROLL_IO".Output[16, 7];
        %Q17.0 := #enabled AND "ROLL_IO".Output[17, 0];
        %Q17.1 := #enabled AND "ROLL_IO".Output[17, 1];
        %Q17.2 := #enabled AND "ROLL_IO".Output[17, 2];
        %Q17.3 := #enabled AND "ROLL_IO".Output[17, 3];
        %Q17.4 := #enabled AND "ROLL_IO".Output[17, 4];
        %Q17.5 := #enabled AND "ROLL_IO".Output[17, 5];
        %Q17.6 := #enabled AND "ROLL_IO".Output[17, 6];
        %Q17.7 := #enabled AND "ROLL_IO".Output[17, 7];
        %Q18.0 := #enabled AND "ROLL_IO".Output[18, 0];
        %Q18.1 := #enabled AND "ROLL_IO".Output[18, 1];
        %Q18.2 := #enabled AND "ROLL_IO".Output[18, 2];
        %Q18.3 := #enabled AND "ROLL_IO".Output[18, 3];
        %Q18.4 := #enabled AND "ROLL_IO".Output[18, 4];
        %Q18.5 := #enabled AND "ROLL_IO".Output[18, 5];
        %Q18.6 := #enabled AND "ROLL_IO".Output[18, 6];
        %Q18.7 := #enabled AND "ROLL_IO".Output[18, 7];
        %Q19.0 := #enabled AND "ROLL_IO".Output[19, 0];
        %Q19.1 := #enabled AND "ROLL_IO".Output[19, 1];
        %Q19.2 := #enabled AND "ROLL_IO".Output[19, 2];
        %Q19.3 := #enabled AND "ROLL_IO".Output[19, 3];
        %Q19.4 := #enabled AND "ROLL_IO".Output[19, 4];
        %Q19.5 := #enabled AND "ROLL_IO".Output[19, 5];
        %Q19.6 := #enabled AND "ROLL_IO".Output[19, 6];
        %Q19.7 := #enabled AND "ROLL_IO".Output[19, 7];
        %Q20.0 := #enabled AND "ROLL_IO".Output[20, 0];
        %Q20.1 := #enabled AND "ROLL_IO".Output[20, 1];
        %Q20.2 := #enabled AND "ROLL_IO".Output[20, 2];
        %Q20.3 := #enabled AND "ROLL_IO".Output[20, 3];
        %Q20.4 := #enabled AND "ROLL_IO".Output[20, 4];
        %Q20.5 := #enabled AND "ROLL_IO".Output[20, 5];
        %Q20.6 := #enabled AND "ROLL_IO".Output[20, 6];
        %Q20.7 := #enabled AND "ROLL_IO".Output[20, 7];
        %Q21.0 := #enabled AND "ROLL_IO".Output[21, 0];
        %Q21.1 := #enabled AND "ROLL_IO".Output[21, 1];
        %Q21.2 := #enabled AND "ROLL_IO".Output[21, 2];
        %Q21.3 := #enabled AND "ROLL_IO".Output[21, 3];
        %Q21.4 := #enabled AND "ROLL_IO".Output[21, 4];
        %Q21.5 := #enabled AND "ROLL_IO".Output[21, 5];
        %Q21.6 := #enabled AND "ROLL_IO".Output[21, 6];
        %Q21.7 := #enabled AND "ROLL_IO".Output[21, 7];
        %Q22.0 := #enabled AND "ROLL_IO".Output[22, 0];
        %Q22.1 := #enabled AND "ROLL_IO".Output[22, 1];
        %Q22.2 := #enabled AND "ROLL_IO".Output[22, 2];
        %Q22.3 := #enabled AND "ROLL_IO".Output[22, 3];
        %Q22.4 := #enabled AND "ROLL_IO".Output[22, 4];
        %Q22.5 := #enabled AND "ROLL_IO".Output[22, 5];
        %Q22.6 := #enabled AND "ROLL_IO".Output[22, 6];
        %Q22.7 := #enabled AND "ROLL_IO".Output[22, 7];
        %Q23.0 := #enabled AND "ROLL_IO".Output[23, 0];
        %Q23.1 := #enabled AND "ROLL_IO".Output[23, 1];
        %Q23.2 := #enabled AND "ROLL_IO".Output[23, 2];
        %Q23.3 := #enabled AND "ROLL_IO".Output[23, 3];
        %Q23.4 := #enabled AND "ROLL_IO".Output[23, 4];
        %Q23.5 := #enabled AND "ROLL_IO".Output[23, 5];
        %Q23.6 := #enabled AND "ROLL_IO".Output[23, 6];
        %Q23.7 := #enabled AND "ROLL_IO".Output[23, 7];
        %Q24.0 := #enabled AND "ROLL_IO".Output[24, 0];
        %Q24.1 := #enabled AND "ROLL_IO".Output[24, 1];
        %Q24.2 := #enabled AND "ROLL_IO".Output[24, 2];
        %Q24.3 := #enabled AND "ROLL_IO".Output[24, 3];
        %Q24.4 := #enabled AND "ROLL_IO".Output[24, 4];
        %Q24.5 := #enabled AND "ROLL_IO".Output[24, 5];
        %Q24.6 := #enabled AND "ROLL_IO".Output[24, 6];
        %Q24.7 := #enabled AND "ROLL_IO".Output[24, 7];
        %Q25.0 := #enabled AND "ROLL_IO".Output[25, 0];
        %Q25.1 := #enabled AND "ROLL_IO".Output[25, 1];
        %Q25.2 := #enabled AND "ROLL_IO".Output[25, 2];
        %Q25.3 := #enabled AND "ROLL_IO".Output[25, 3];
        %Q25.4 := #enabled AND "ROLL_IO".Output[25, 4];
        %Q25.5 := #enabled AND "ROLL_IO".Output[25, 5];
        %Q25.6 := #enabled AND "ROLL_IO".Output[25, 6];
        %Q25.7 := #enabled AND "ROLL_IO".Output[25, 7];
    END_IF;
END_FUNCTION

FUNCTION "ROLL_HmiExchange" : Void
{ S7_Optimized_Access := 'TRUE' }
VERSION : 0.1
VAR_INPUT
    DeltaMs : LReal;
END_VAR
VAR_TEMP
    b : Int;
    bit : Int;
    n : Int;
    fieldIndex : Int;
    index : Int;
    raw : Word;
    base : DInt;
    count : DInt;
    recipe : Array[0..41] of Word;
END_VAR
BEGIN
    // Called at the end of the scan, like the former OP15 functions in OB1.
    "ROLL_IO".HmiElapsedMs := "ROLL_IO".HmiElapsedMs + #DeltaMs;
    IF "ROLL_HMI".Heartbeat <> "ROLL_IO".HmiLastHeartbeat THEN
        "ROLL_IO".HmiLastHeartbeat := "ROLL_HMI".Heartbeat;
        "ROLL_IO".HmiElapsedMs := 0.0;
        "ROLL_HMI".Connected := TRUE;
    END_IF;
    IF "ROLL_IO".HmiElapsedMs >= 1500.0 THEN "ROLL_HMI".Connected := FALSE; END_IF;
    "ROLL_State".M[190, 5] := "ROLL_HMI".Connected AND "ROLL_HMI".GroundHeld;
    "ROLL_State".M[190, 6] := "ROLL_HMI".Connected AND "ROLL_HMI".WorkHeld;
    "ROLL_State".M[190, 3] := ("ROLL_State".M[190, 5] OR "ROLL_State".M[190, 6]) AND NOT "ROLL_State".M[190, 4];
    "ROLL_State".M[190, 4] := "ROLL_State".M[190, 5] OR "ROLL_State".M[190, 6];
    "ROLL_State".M[191, 0] := FALSE;
    IF ("ROLL_HMI".ManualFunction >= 0) AND ("ROLL_HMI".ManualFunction <= 255) AND "ROLL_HMI".Connected THEN
        "ROLL_SetMWord"(FirstByte := 238, Value := INT_TO_WORD("ROLL_HMI".ManualFunction));
    ELSE
        "ROLL_SetMWord"(FirstByte := 238, Value := W#16#00FF);
    END_IF;
    FOR #n := 0 TO 7 DO
        "ROLL_State".M[192, #n] := "ROLL_HMI".Connected AND "ROLL_HMI".KeyF[#n + 1];
        "ROLL_State".M[193, #n] := "ROLL_HMI".Connected AND "ROLL_HMI".KeyF[#n + 9];
    END_FOR;

    // Request/acknowledgement counters prevent partial edits on every scan.
    // Command 1 loads the retained program; command 2 saves the displayed values.
    IF "ROLL_HMI".RecipeRequest <> "ROLL_HMI".RecipeAck THEN
        "ROLL_HMI".RecipeError := 0;
        IF NOT "ROLL_HMI".Connected THEN
            "ROLL_HMI".RecipeError := 8;
        ELSIF ("ROLL_HMI".SelectedProgram < 1) OR ("ROLL_HMI".SelectedProgram > 2) THEN
            "ROLL_HMI".RecipeError := 1;
        ELSIF NOT "ROLL_IO".Input[0, 1] THEN
            "ROLL_HMI".RecipeError := 2; // requires manual operating mode
        ELSIF ("ROLL_HMI".RecipeCommand <> 1) AND ("ROLL_HMI".RecipeCommand <> 2) THEN
            "ROLL_HMI".RecipeError := 3;
        ELSE
            FOR #n := 0 TO 41 DO
                IF "ROLL_HMI".SelectedProgram = 1 THEN #recipe[#n] := "ROLL_Recipe1".DW[#n];
                ELSE #recipe[#n] := "ROLL_Recipe2".DW[#n]; END_IF;
            END_FOR;
            IF "ROLL_HMI".RecipeCommand = 2 THEN
                #recipe[5] := "ROLL_EncodeSeconds"(Seconds := "ROLL_HMI".Dwell1Seconds);
                #recipe[9] := "ROLL_EncodeSeconds"(Seconds := "ROLL_HMI".Drain1Seconds);
                #recipe[17] := "ROLL_EncodeSeconds"(Seconds := "ROLL_HMI".Dwell2Seconds);
                #recipe[21] := "ROLL_EncodeSeconds"(Seconds := "ROLL_HMI".Drain2Seconds);
                #recipe[25] := "ROLL_EncodeSeconds"(Seconds := "ROLL_HMI".Dwell3Seconds);
                #recipe[29] := "ROLL_EncodeSeconds"(Seconds := "ROLL_HMI".Drain3Seconds);
                #recipe[33] := "ROLL_EncodeSeconds"(Seconds := "ROLL_HMI".Dry4Seconds);
                FOR #n := 0 TO 6 DO
                    CASE #n OF
                        0: #fieldIndex := 5; 1: #fieldIndex := 9; 2: #fieldIndex := 17;
                        3: #fieldIndex := 21; 4: #fieldIndex := 25; 5: #fieldIndex := 29;
                        6: #fieldIndex := 33;
                    END_CASE;
                    IF #recipe[#fieldIndex] = W#16#FFFF THEN "ROLL_HMI".RecipeError := 4; END_IF;
                END_FOR;
                IF ("ROLL_HMI".BasketMotion < 0) OR ("ROLL_HMI".BasketMotion > 4) THEN "ROLL_HMI".RecipeError := 5; END_IF;
                #recipe[37] := INT_TO_WORD("ROLL_HMI".BasketMotion);
                #recipe[13] := W#16#0000;
                IF "ROLL_HMI".Ultrasound1 THEN #recipe[13] := W#16#0001; END_IF;
                #recipe[41] := W#16#0000;
                IF "ROLL_HMI".BathLift THEN #recipe[41] := W#16#0001; END_IF;
            END_IF;
            IF "ROLL_HMI".RecipeError = 0 THEN
                FOR #n := 0 TO 41 DO
                    "ROLL_DB205".DW[#n] := #recipe[#n];
                    IF "ROLL_HMI".RecipeCommand = 2 THEN
                        IF "ROLL_HMI".SelectedProgram = 1 THEN "ROLL_Recipe1".DW[#n] := #recipe[#n];
                        ELSE "ROLL_Recipe2".DW[#n] := #recipe[#n]; END_IF;
                    END_IF;
                END_FOR;
                "ROLL_State".CurrentProgram := "ROLL_HMI".SelectedProgram;
                "ROLL_ShowRecipe"();
                "ROLL_State".M[190, 1] := TRUE;
                "ROLL_State".M[190, 2] := FALSE;
                "ROLL_State".M[191, 4] := TRUE;
                "ROLL_FB90"();
            END_IF;
        END_IF;
        "ROLL_HMI".RecipeAck := "ROLL_HMI".RecipeRequest;
    END_IF;

    IF "ROLL_HMI".ParameterRequest <> "ROLL_HMI".ParameterAck THEN
        "ROLL_HMI".ParameterError := 0;
        #index := "ROLL_HMI".ParameterIndex;
        #raw := W#16#FFFF;
        IF NOT "ROLL_HMI".Connected THEN "ROLL_HMI".ParameterError := 8;
        ELSIF (#index < 0) OR (#index > 127) THEN "ROLL_HMI".ParameterError := 1;
        ELSIF NOT "ROLL_IO".Input[0, 1] THEN "ROLL_HMI".ParameterError := 2;
        ELSIF ("ROLL_HMI".ParameterDb <> 15) AND ("ROLL_HMI".ParameterDb <> 19) THEN "ROLL_HMI".ParameterError := 3;
        ELSE
            #raw := "ROLL_GetDW"(DbNumber := "ROLL_HMI".ParameterDb, Index := #index);
            IF #raw = W#16#FFFF THEN "ROLL_HMI".ParameterError := 4;
            ELSE
                #base := 1;
                IF "ROLL_HMI".ParameterDb = 15 THEN
                    CASE WORD_TO_INT(SHR(IN := #raw AND W#16#F000, N := 12)) OF
                        0: #base := 10; 1: #base := 100; 2: #base := 1000; 3: #base := 10000;
                        ELSE #base := 0;
                    END_CASE;
                END_IF;
                IF #base = 0 THEN "ROLL_HMI".ParameterError := 5;
                ELSIF ("ROLL_HMI".ParameterValue < 0) OR (("ROLL_HMI".ParameterValue MOD #base) <> 0) THEN "ROLL_HMI".ParameterError := 6;
                ELSE
                    #count := "ROLL_HMI".ParameterValue / #base;
                    IF #count > 999 THEN "ROLL_HMI".ParameterError := 7;
                    ELSE
                        #raw := (#raw AND W#16#F000) OR SHL(IN := DINT_TO_WORD(#count / 100), N := 8)
                            OR SHL(IN := DINT_TO_WORD((#count / 10) MOD 10), N := 4) OR DINT_TO_WORD(#count MOD 10);
                        IF "ROLL_HMI".ParameterDb = 15 THEN "ROLL_DB15".DW[#index] := #raw;
                        ELSE "ROLL_DB19".DW[#index] := #raw; END_IF;
                    END_IF;
                END_IF;
            END_IF;
        END_IF;
        "ROLL_HMI".ParameterAck := "ROLL_HMI".ParameterRequest;
    END_IF;
    "ROLL_HMI".ParameterSlotPresent := FALSE;
    "ROLL_HMI".ParameterCurrentValue := 0;
    #index := "ROLL_HMI".ParameterIndex;
    IF (#index >= 0) AND (#index <= 127) AND (("ROLL_HMI".ParameterDb = 15) OR ("ROLL_HMI".ParameterDb = 19)) THEN
        #raw := "ROLL_GetDW"(DbNumber := "ROLL_HMI".ParameterDb, Index := #index);
        IF #raw <> W#16#FFFF THEN
            #count := INT_TO_DINT("ROLL_DecodeBCD"(Value := #raw));
            #base := 1;
            IF "ROLL_HMI".ParameterDb = 15 THEN
                CASE WORD_TO_INT(SHR(IN := #raw AND W#16#F000, N := 12)) OF
                    0: #base := 10; 1: #base := 100; 2: #base := 1000; 3: #base := 10000;
                    ELSE #base := 0;
                END_CASE;
            END_IF;
            IF (#count >= 0) AND (#base > 0) THEN
                "ROLL_HMI".ParameterSlotPresent := TRUE;
                "ROLL_HMI".ParameterCurrentValue := #count * #base;
            END_IF;
        END_IF;
    END_IF;
    IF WORD_TO_INT("ROLL_GetM"(FirstByte := 239, Width := 8)) <> 255 THEN
        "ROLL_PB18"();
    ELSE
        "ROLL_SetMWord"(FirstByte := 250, Value := W#16#0000);
        "ROLL_SetMWord"(FirstByte := 252, Value := W#16#0000);
    END_IF;
    "ROLL_HMI".ProcessTimer1Units := WORD_TO_INT("ROLL_TimerValue"(Number := 1));
    "ROLL_HMI".ProcessTimer2Units := WORD_TO_INT("ROLL_TimerValue"(Number := 2));
    FOR #b := 0 TO 255 DO
        FOR #bit := 0 TO 7 DO "ROLL_HMI".StatusM[#b, #bit] := "ROLL_State".M[#b, #bit]; END_FOR;
    END_FOR;
    FOR #b := 16 TO 25 DO
        FOR #bit := 0 TO 7 DO "ROLL_HMI".LogicalOutputs[#b, #bit] := "ROLL_IO".Output[#b, #bit]; END_FOR;
    END_FOR;
END_FUNCTION

FUNCTION "ROLL_Cycle" : Void
{ S7_Optimized_Access := 'TRUE' }
VERSION : 0.1
VAR_TEMP
    delta : LReal;
END_VAR
BEGIN
    #delta := RUNTIME("ROLL_IO".RuntimeMemory) * 1000.0;
    IF "ROLL_IO".FirstCycle THEN
        #delta := 0.0;
        "ROLL_IO".FirstCycle := FALSE;
    END_IF;
    "ROLL_ReadInputs"();
    "ROLL_AdvanceTime"(DeltaMs := #delta);
    // Exact OB1 order for the process blocks; startup DB creation is replaced.
    IF NOT "ROLL_State".M[0, 2] THEN "ROLL_State".M[0, 1] := FALSE; END_IF;
    IF "ROLL_State".M[0, 1] THEN "ROLL_State".M[0, 7] := TRUE; END_IF;
    "ROLL_State".M[0, 5] := NOT "ROLL_State".M[0, 5];
    IF "ROLL_State".M[3, 2] THEN "ROLL_State".M[3, 3] := TRUE; END_IF;
    IF "ROLL_IO".Input[0, 2] THEN "ROLL_State".M[3, 3] := FALSE; END_IF;
    "ROLL_State".M[3, 2] := "ROLL_IO".Input[0, 1] AND NOT "ROLL_State".M[0, 1];
    "ROLL_PB2"();
    IF "ROLL_State".M[0, 7] THEN "ROLL_State".M[0, 7] := FALSE; END_IF;
    "ROLL_PB3"();
    "ROLL_PB4"();
    "ROLL_PB19"();
    "ROLL_PB21"();
    "ROLL_PB50"();
    "ROLL_PB51"();
    "ROLL_PB52"();
    IF NOT "ROLL_State".M[3, 3] THEN "ROLL_PB8"(); END_IF;
    IF NOT "ROLL_State".M[3, 3] THEN "ROLL_PB9"(); END_IF;
    IF NOT "ROLL_State".M[3, 3] THEN "ROLL_PB10"(); END_IF;
    IF NOT "ROLL_State".M[3, 3] THEN "ROLL_PB14"(); END_IF;
    IF "ROLL_State".M[3, 3] THEN "ROLL_PB16"(); END_IF;
    "ROLL_PB7"();
    "ROLL_PB13"();
    "ROLL_PB15"();
    "ROLL_PB17"();
    "ROLL_PB20"();
    "ROLL_PB23"();
    "ROLL_PB24"();
    "ROLL_PB25"();
    "ROLL_FB111"();
    "ROLL_HmiExchange"(DeltaMs := #delta);
    "ROLL_WriteOutputs"();
END_FUNCTION

ORGANIZATION_BLOCK OB100
{ S7_Optimized_Access := 'TRUE' }
VERSION : 0.1
VAR_TEMP
    n : Int;
END_VAR
BEGIN
    // RE plus RS120 bit 3: all M retained. Default T/Z 0..63 retained.
    FOR #n := 64 TO 127 DO
        "ROLL_State".S5Timers[#n].RemainingMs := 0.0;
        "ROLL_State".S5Timers[#n].BaseMs := 0;
        "ROLL_State".S5Timers[#n].Mode := 0;
        "ROLL_State".S5Timers[#n].Q := FALSE;
        "ROLL_State".S5Timers[#n].Previous := FALSE;
        "ROLL_State".S5Counters[#n].Value := 0;
        "ROLL_State".S5Counters[#n].SetPrevious := FALSE;
        "ROLL_State".S5Counters[#n].UpPrevious := FALSE;
        "ROLL_State".S5Counters[#n].DownPrevious := FALSE;
    END_FOR;
    "ROLL_IO".FirstCycle := TRUE;
    "ROLL_IO".ClockMs := 0.0;
    "ROLL_IO".RuntimeMemory := 0.0;
    "ROLL_IO".PhysicalOutputsEnabled := FALSE;
    "ROLL_HMI".Connected := FALSE;
    "ROLL_State".M[0, 1] := TRUE;
    "ROLL_State".M[0, 2] := TRUE;
    "ROLL_State".M[191, 0] := TRUE;
    "ROLL_State".M[190, 5] := FALSE;
    "ROLL_State".M[190, 6] := FALSE;
    "ROLL_State".M[190, 1] := TRUE;
    "ROLL_State".M[191, 4] := TRUE;
    "ROLL_FB90"();
    "ROLL_ShowRecipe"();
END_ORGANIZATION_BLOCK

ORGANIZATION_BLOCK OB1
{ S7_Optimized_Access := 'TRUE' }
VERSION : 0.1
BEGIN
    "ROLL_Cycle"();
END_ORGANIZATION_BLOCK
